(* IEC 61131-3 sources: codesys-to-s7/tests/corpus/C2S7-SEM-MUX/neg, 1 file *)

(* ---- input.st ---- *)
FUNCTION_BLOCK FB_Case
VAR
    a : INT;
    b : INT;
    i : INT;
    d : DINT;
    r : REAL;
    x : BOOL;
    y : BOOL;
    s : STRING(80);
    w : WORD;
    t : TIME;
END_VAR
i := SEL(x, 1, 2);
END_FUNCTION_BLOCK
